(* Communication structure from plc to drive *)

TYPE ST_PLCTOBECKHOFFDRIVE :
STRUCT
		wPO1ControlWord						:WORD;
END_STRUCT
END_TYPE

(* stored: Version 1.1.0.1, ProductVersion 3.1.4024.15
   DUT ST_PLCTOBECKHOFFDRIVE: Id {01b5c534-2c26-49ce-8466-9462d3b5eba7} *)
